{attribute 'qualified_only'}
{attribute 'strict'}
{attribute 'to_string'}
TYPE E_LineState :
(
    Stopped      := 0,
    Filling      := 10,
    Transferring := 20,
    Faulted      := 900
);
END_TYPE

(* stored: Version 1.1.0.1
   DUT E_LineState: Id {56a82c92-05b6-4f4e-9811-e9a859d97f8b} *)
